Fanuc KAREL source: kt00212.KL

-- PROVISIONAL review KL for V940-1; original PC SHA256 81a7c44bc666b1bb721210bad6b797378683cc4acab3aed75838bbf299bbd5bf
-- Incomplete behavior may be omitted. Consult companion uncertainty JSON. Do not deploy.
PROGRAM KT00212
%NOLOCKGROUP
VAR
  I2 : INTEGER
  OUT : INTEGER
-- UNRESOLVED_DECL Y1 type=002018
BEGIN
  -- V9_ZERO_TABLE_METADATA_HINT layout=0001; no indexed target words; source/name/runtime held
  -- UNRESOLVED_PC offsets 5-19; opcodes 2E,22,9D,33,B2
  -- UNRESOLVED_PC offsets 24-35; opcodes 2E,23
  -- UNRESOLVED_PC offsets 40-62; opcodes 22,9D,33,B1,21,46,23
  -- UNRESOLVED_PC offsets 67-71; opcodes 7F
END KT00212
